Fanuc KAREL source: kd00045.KL

-- PROVISIONAL review KL for V940-1; original PC SHA256 a1996fe47cd37e1b99638785196df67873e3dca7f7c603beb26e81fbaa66ca19
-- Incomplete behavior may be omitted. Consult companion uncertainty JSON. Do not deploy.
PROGRAM KD00045
%NOLOCKGROUP
VAR
  I : INTEGER
  J : INTEGER
  B : BOOLEAN
  R : REAL
  S : STRING[80]
-- UNRESOLVED_DECL P type=000101
BEGIN
  -- V9_ZERO_TABLE_METADATA_HINT layout=0001; no indexed target words; source/name/runtime held
  -- UNRESOLVED_PC offsets 5-24; opcodes 01,22,1C,06,82,0B
  -- UNRESOLVED_PC offsets 29-33; opcodes 7F
END KD00045
